// HMI -> PLC: gate requests (Tap). A request only; unlocking stays with the safety logic.
TYPE ST_HMI_GateCommand :
STRUCT
    bRequestAccess : BOOL;
    bReset : BOOL;
END_STRUCT
END_TYPE

(* stored: Version 1.1.0.1
   DUT ST_HMI_GateCommand: Id {2d9fcf5c-3e7a-4c3d-a199-6e13dd43daba} *)
